Fanuc KAREL source: KT00073.KL

PROGRAM KT00073
%NOLOCKGROUP
VAR
  R1: REAL
  I2: INTEGER
  OUT: INTEGER
BEGIN
  R1 = 2.0
    I2 = 3
  OUT = R1 * I2
END KT00073
